TYPE ST_AlarmProperties_1 :
STRUCT
	bActive				:BOOL;				(* Alarm on *)
	{attribute 'hide'} 
	dtDateTime			:DATE_AND_TIME ;	(* Alarm time stamp *)
	{attribute 'hide'} 
	enType				:ET_AlarmType;		(* Alarm type *)
	dnCode				:DINT;				(* Alarm code *)
END_STRUCT
END_TYPE

(* stored: Version 1.1.0.1, ProductVersion 3.1.4024.15
   DUT ST_AlarmProperties_1: Id {f2ac693c-7322-476b-ae3d-f84e1f585277} *)
